                num nValue[3]
            mdesc mMdesc = {accel=25, vel=50, leave=1}
            num nActionIndex = 8
            num nDelay
            num nMoveType = 1
            num nPercentage
            num nSigValue = 1
        pointRx pPointRx[2] = {x=594.549716, y=30.77075, z=284.629716, rx=-40.404847, ry=94.502137, rz=40.914396, shoulder=lefty, elbow=epositive, wrist=wnegative}
        string sID
      [17]
        bool bMarked
        jointRx jJointRx = {j1=-1.639045, j2=12.402747, j3=111.595585, j4=2.517874, j5=-30.594648, j6=-1.669011}
        pointRx pInter
        paraItem pParaItem
          [0]
            bool bSafePoint
            ifItem iIfItem
              [0]
                bool bANDOR[2]
                num nSigIndex[3]
                num nSigType[3]
                num nValue[3]
            mdesc mMdesc
            num nActionIndex = 10
            num nDelay = 5
            num nMoveType = 4
            num nPercentage
            num nSigValue
        pointRx pPointRx[2] = {x=594.549819, y=30.770866, z=171.45682, rx=-40.410864, ry=94.502866, rz=40.920287, shoulder=lefty, elbow=epositive, wrist=wnegative}
        string sID
      [18]
        bool bMarked
        jointRx jJointRx = {j1=-1.639045, j2=12.402747, j3=111.595585, j4=2.517874, j5=-30.594648, j6=-1.669011}
        pointRx pInter
        paraItem pParaItem
          [0]
            bool bSafePoint
            ifItem iIfItem
              [0]
                bool bANDOR[2]
                num nSigIndex[3]
                num nSigType[3]
                num nValue[3]
            mdesc mMdesc
            num nActionIndex = 10
            num nDelay = 0.5
            num nMoveType = 7
            num nPercentage
            num nSigValue
        pointRx pPointRx[2] = {x=594.549819, y=30.770866, z=171.45682, rx=-40.410864, ry=94.502866, rz=40.920287, shoulder=lefty, elbow=epositive, wrist=wnegative}
        string sID
      [19]
        bool bMarked
        jointRx jJointRx = {j1=-1.639045, j2=12.402747, j3=111.595585, j4=2.517874, j5=-30.594648, j6=-1.669011}
        pointRx pInter
        paraItem pParaItem
          [0]
            bool bSafePoint
            ifItem iIfItem
              [0]
                bool bANDOR[2]
                num nSigIndex[3]
                num nSigType[3]
                num nValue[3]
            mdesc mMdesc
            num nActionIndex = 9
            num nDelay = 5
            num nMoveType = 3
            num nPercentage
            num nSigValue = 1
        pointRx pPointRx[2] = {x=594.549819, y=30.770866, z=171.45682, rx=-40.410864, ry=94.502866, rz=40.920287, shoulder=lefty, elbow=epositive, wrist=wnegative}
        string sID
      [20]
        bool bMarked
        jointRx jJointRx = {j1=-1.639045, j2=12.402747, j3=111.595585, j4=2.517874, j5=-30.594648, j6=-1.669011}
        pointRx pInter
        paraItem pParaItem
          [0]
            bool bSafePoint
            ifItem iIfItem
              [0]
                bool bANDOR[2]
                num nSigIndex[3]
                num nSigType[3]
                num nValue[3]
            mdesc mMdesc
            num nActionIndex = 9
            num nDelay = 5
            num nMoveType
            num nPercentage
            num nSigValue = 1
        pointRx pPointRx[2] = {x=594.549819, y=30.770866, z=171.45682, rx=-40.410864, ry=94.502866, rz=40.920287, shoulder=lefty, elbow=epositive, wrist=wnegative}
        string sID
      [21]
        bool bMarked
        jointRx jJointRx = {j1=-1.639045, j2=12.402747, j3=111.595585, j4=2.517874, j5=-30.594648, j6=-1.669011}
        pointRx pInter
        paraItem pParaItem
          [0]
            bool bSafePoint
            ifItem iIfItem
              [0]
                bool bANDOR[2]
                num nSigIndex[3]
                num nSigType[3]
                num nValue[3]
            mdesc mMdesc
            num nActionIndex = 9
            num nDelay = 5
            num nMoveType = 1
            num nPercentage
            num nSigValue = 1
        pointRx pPointRx[2] = {x=594.549819, y=30.770866, z=171.45682, rx=-40.410864, ry=94.502866, rz=40.920287, shoulder=lefty, elbow=epositive, wrist=wnegative}
        string sID
      [22]
        bool bMarked
        jointRx jJointRx = {j1=-1.639045, j2=12.402747, j3=111.595585, j4=2.517874, j5=-30.594648, j6=-1.669011}
        pointRx pInter
        paraItem pParaItem
          [0]
            bool bSafePoint
            ifItem iIfItem
              [0]
                bool bANDOR[2]
                num nSigIndex[3]
                num nSigType[3]
                num nValue[3]
            mdesc mMdesc
            num nActionIndex = 1
            num nDelay = 5
            num nMoveType = 6
            num nPercentage
            num nSigValue = 3
        pointRx pPointRx[2] = {x=594.549819, y=30.770866, z=171.45682, rx=-40.410864, ry=94.502866, rz=40.920287, shoulder=lefty, elbow=epositive, wrist=wnegative}
        string sID
      [23]
        bool bMarked
        jointRx jJointRx = {j1=-1.639045, j2=12.402747, j3=111.595585, j4=2.517874, j5=-30.594648, j6=-1.669011}
        pointRx pInter
        paraItem pParaItem
          [0]
            bool bSafePoint
            ifItem iIfItem
              [0]
                bool bANDOR[2]
                num nSigIndex[3]
                num nSigType[3]
                num nValue[3]
            mdesc mMdesc
            num nActionIndex = 1
            num nDelay = 5
            num nMoveType = 5
            num nPercentage
            num nSigValue = 3
        pointRx pPointRx[2] = {x=594.549819, y=30.770866, z=171.45682, rx=-40.410864, ry=94.502866, rz=40.920287, shoulder=lefty, elbow=epositive, wrist=wnegative}
        string sID
      [24]
        bool bMarked
        jointRx jJointRx = {j1=-1.639045, j2=12.402747, j3=111.595585, j4=2.517874, j5=-30.594648, j6=-1.669011}
        pointRx pInter
        paraItem pParaItem
          [0]
            bool bSafePoint
            ifItem iIfItem
              [0]
                bool bANDOR[2]
                num nSigIndex[3]
                num nSigType[3]
                num nValue[3]
            mdesc mMdesc
            num nActionIndex = 10
            num nDelay
            num nMoveType = 4
            num nPercentage
            num nSigValue = 1
        pointRx pPointRx[2] = {x=594.549819, y=30.770866, z=171.45682, rx=-40.410864, ry=94.502866, rz=40.920287, shoulder=lefty, elbow=epositive, wrist=wnegative}
        string sID
      [25]
        bool bMarked
        jointRx jJointRx = {j1=-1.639045, j2=12.402747, j3=111.595585, j4=2.517874, j5=-30.594648, j6=-1.669011}
        pointRx pInter
        paraItem pParaItem
          [0]
            bool bSafePoint
            ifItem iIfItem
              [0]
                bool bANDOR[2]
                num nSigIndex[3]
                num nSigType[3]
                num nValue[3]
            mdesc mMdesc
            num nActionIndex = 8
            num nDelay
            num nMoveType = 3
            num nPercentage
            num nSigValue = 1
        pointRx pPointRx[2] = {x=594.549819, y=30.770866, z=171.45682, rx=-40.410864, ry=94.502866, rz=40.920287, shoulder=lefty, elbow=epositive, wrist=wnegative}
        string sID
      [26]
        bool bMarked
        jointRx jJointRx = {j1=-1.639134, j2=22.193742, j3=116.03978, j4=1.817031, j5=-44.819098, j6=-0.790246}
        pointRx pInter
        paraItem pParaItem
          [0]
            bool bSafePoint
            ifItem iIfItem
              [0]
                bool bANDOR[2]
                num nSigIndex[3]
                num nSigType[3]
                num nValue[3]
            mdesc mMdesc = {accel=25, vel=50, leave=1}
            num nActionIndex = 8
            num nDelay
            num nMoveType = 1
            num nPercentage
            num nSigValue = 1
        pointRx pPointRx[2] = {x=594.549757, y=30.770873, z=70.540177, rx=-40.399083, ry=94.503271, rz=40.908669, shoulder=lefty, elbow=epositive, wrist=wnegative}
        string sID
      [27]
        bool bMarked
        jointRx jJointRx = {j1=-1.639045, j2=12.402747, j3=111.595585, j4=2.517874, j5=-30.594648, j6=-1.669011}
        pointRx pInter
        paraItem pParaItem
          [0]
            bool bSafePoint
            ifItem iIfItem
              [0]
                bool bANDOR[2]
                num nSigIndex[3]
                num nSigType[3]
                num nValue[3]
            mdesc mMdesc
            num nActionIndex = 10
            num nDelay = 5
            num nMoveType = 4
            num nPercentage
            num nSigValue
        pointRx pPointRx[2] = {x=594.549819, y=30.770866, z=171.45682, rx=-40.410864, ry=94.502866, rz=40.920287, shoulder=lefty, elbow=epositive, wrist=wnegative}
        string sID
      [28]
        bool bMarked
        jointRx jJointRx = {j1=-1.639045, j2=12.402747, j3=111.595585, j4=2.517874, j5=-30.594648, j6=-1.669011}
        pointRx pInter
        paraItem pParaItem
          [0]
            bool bSafePoint
            ifItem iIfItem
              [0]
                bool bANDOR[2]
                num nSigIndex[3]
                num nSigType[3]
                num nValue[3]
            mdesc mMdesc
            num nActionIndex = 10
            num nDelay = 0.5
            num nMoveType = 7
            num nPercentage
            num nSigValue
        pointRx pPointRx[2] = {x=594.549819, y=30.770866, z=171.45682, rx=-40.410864, ry=94.502866, rz=40.920287, shoulder=lefty, elbow=epositive, wrist=wnegative}
        string sID
      [29]
        bool bMarked
        jointRx jJointRx = {j1=-1.639045, j2=12.402747, j3=111.595585, j4=2.517874, j5=-30.594648, j6=-1.669011}
        pointRx pInter
        paraItem pParaItem
          [0]
            bool bSafePoint
            ifItem iIfItem
              [0]
                bool bANDOR[2]
                num nSigIndex[3]
                num nSigType[3]
                num nValue[3]
            mdesc mMdesc
            num nActionIndex = 9
            num nDelay = 5
            num nMoveType = 3
            num nPercentage
            num nSigValue = 1
        pointRx pPointRx[2] = {x=594.549819, y=30.770866, z=171.45682, rx=-40.410864, ry=94.502866, rz=40.920287, shoulder=lefty, elbow=epositive, wrist=wnegative}
        string sID
      [30]
        bool bMarked
        jointRx jJointRx = {j1=-1.639045, j2=12.402747, j3=111.595585, j4=2.517874, j5=-30.594648, j6=-1.669011}
        pointRx pInter
        paraItem pParaItem
          [0]
            bool bSafePoint
            ifItem iIfItem
              [0]
                bool bANDOR[2]
                num nSigIndex[3]
                num nSigType[3]
                num nValue[3]
            mdesc mMdesc
            num nActionIndex = 1
            num nDelay = 5
            num nMoveType = 6
            num nPercentage
            num nSigValue
        pointRx pPointRx[2] = {x=594.549819, y=30.770866, z=171.45682, rx=-40.410864, ry=94.502866, rz=40.920287, shoulder=lefty, elbow=epositive, wrist=wnegative}
        string sID
      [31]
        bool bMarked
        jointRx jJointRx = {j1=-1.639045, j2=12.402747, j3=111.595585, j4=2.517874, j5=-30.594648, j6=-1.669011}
        pointRx pInter
        paraItem pParaItem
          [0]
            bool bSafePoint
            ifItem iIfItem
              [0]
                bool bANDOR[2]
                num nSigIndex[3]
                num nSigType[3]
                num nValue[3]
            mdesc mMdesc
            num nActionIndex = 1
            num nDelay = 5
            num nMoveType = 5
            num nPercentage
            num nSigValue
        pointRx pPointRx[2] = {x=594.549819, y=30.770866, z=171.45682, rx=-40.410864, ry=94.502866, rz=40.920287, shoulder=lefty, elbow=epositive, wrist=wnegative}
        string sID
      [32]
        bool bMarked
        jointRx jJointRx = {j1=-6.64887, j2=-3.725236, j3=129.0447824, j4=-6.346176, j5=-34.648626, j6=4.794545}
        pointRx pInter
        paraItem pParaItem
          [0]
            bool bSafePoint
            ifItem iIfItem
              [0]
                bool bANDOR[2]
                num nSigIndex[3]
                num nSigType[3]
                num nValue[3]
            mdesc mMdesc
            num nActionIndex = 1
            num nDelay = 5
            num nMoveType
            num nPercentage
            num nSigValue
        pointRx pPointRx[2] = {x=472.316216, y=1.60837, z=176.938996, rx=-74.680282, ry=93.157396, rz=74.321891, shoulder=lefty, elbow=epositive, wrist=wnegative}
        string sID
      [33]
        bool bMarked
        jointRx jJointRx = {j1=-1.639045, j2=12.402747, j3=111.595585, j4=2.517874, j5=-30.594648, j6=-1.669011}
        pointRx pInter
        paraItem pParaItem
          [0]
            bool bSafePoint
            ifItem iIfItem
              [0]
                bool bANDOR[2]
                num nSigIndex[3]
                num nSigType[3]
                num nValue[3]
            mdesc mMdesc
            num nActionIndex = 11
            num nDelay = 5
            num nMoveType = 4
            num nPercentage
            num nSigValue = 1
        pointRx pPointRx[2] = {x=594.549819, y=30.770866, z=171.45682, rx=-40.410864, ry=94.502866, rz=40.920287, shoulder=lefty, elbow=epositive, wrist=wnegative}
        string sID
      [34]
        bool bMarked
        jointRx jJointRx = {j1=-1.639045, j2=12.402747, j3=111.595585, j4=2.517874, j5=-30.594648, j6=-1.669011}
        pointRx pInter
        paraItem pParaItem
          [0]
            bool bSafePoint
            ifItem iIfItem
              [0]
                bool bANDOR[2]
                num nSigIndex[3]
                num nSigType[3]
                num nValue[3]
            mdesc mMdesc
            num nActionIndex = 10
            num nDelay = 5
            num nMoveType = 3
            num nPercentage
            num nSigValue
        pointRx pPointRx[2] = {x=594.549819, y=30.770866, z=171.45682, rx=-40.410864, ry=94.502866, rz=40.920287, shoulder=lefty, elbow=epositive, wrist=wnegative}
        string sID
      [35]
        bool bMarked
        jointRx jJointRx = {j1=-1.639045, j2=12.402747, j3=111.595585, j4=2.517874, j5=-30.594648, j6=-1.669011}
        pointRx pInter
        paraItem pParaItem
          [0]
            bool bSafePoint
            ifItem iIfItem
              [0]
                bool bANDOR[2]
                num nSigIndex[3]
                num nSigType[3]
                num nValue[3]
            mdesc mMdesc
            num nActionIndex = 9
            num nDelay = 5
            num nMoveType = 4
            num nPercentage
            num nSigValue
        pointRx pPointRx[2] = {x=594.549819, y=30.770866, z=171.45682, rx=-40.410864, ry=94.502866, rz=40.920287, shoulder=lefty, elbow=epositive, wrist=wnegative}
        string sID
      [36]
        bool bMarked
        jointRx jJointRx = {j1=-1.639045, j2=12.402747, j3=111.595585, j4=2.517874, j5=-30.594648, j6=-1.669011}
        pointRx pInter
        paraItem pParaItem
          [0]
            bool bSafePoint
            ifItem iIfItem
              [0]
                bool bANDOR[2]
                num nSigIndex[3]
                num nSigType[3]
                num nValue[3]
            mdesc mMdesc
            num nActionIndex = 11
            num nDelay = 5
            num nMoveType = 4
            num nPercentage
            num nSigValue
        pointRx pPointRx[2] = {x=594.549819, y=30.770866, z=171.45682, rx=-40.410864, ry=94.502866, rz=40.920287, shoulder=lefty, elbow=epositive, wrist=wnegative}
        string sID
    string sID
  [03 543-7-0741]
    num nFrameIndex
    num nMoveID
    num nToolIndex
    pointItem pPointItem[45]
      [0]
        bool bMarked
        jointRx jJointRx = {j1=-2.594987, j2=-12.391258, j3=136.392534, j4=0.644488, j5=-30.575639, j6=-0.113504}
        pointRx pInter
        paraItem pParaItem
          [0]
            bool bSafePoint
            ifItem iIfItem
              [0]
                bool bANDOR[2]
                num nSigIndex[3]
                num nSigType[3]
                num nValue[3]
            mdesc mMdesc
            num nActionIndex = 11
            num nDelay
            num nMoveType = 4
            num nPercentage
            num nSigValue
        pointRx pPointRx[2] = {x=412.772469, y=30.77087, z=171.456836, rx=-40.418431, ry=94.503508, rz=40.927655, shoulder=lefty, elbow=epositive, wrist=wnegative}
        string sID
      [1]
        bool bMarked
        jointRx jJointRx = {j1=-2.594987, j2=-12.391258, j3=136.392534, j4=0.644488, j5=-30.575639, j6=-0.113504}
        pointRx pInter
        paraItem pParaItem
          [0]
            bool bSafePoint
            ifItem iIfItem
              [0]
                bool bANDOR[2]
                num nSigIndex[3]
                num nSigType[3]
                num nValue[3]
            mdesc mMdesc
            num nActionIndex = 9
            num nDelay
            num nMoveType = 4
            num nPercentage
            num nSigValue = 1
        pointRx pPointRx[2] = {x=412.772469, y=30.77087, z=171.456836, rx=-40.418431, ry=94.503508, rz=40.927655, shoulder=lefty, elbow=epositive, wrist=wnegative}
        string sID
      [2]
        bool bMarked
        jointRx jJointRx = {j1=-6.652009, j2=-3.724795, j3=129.0452396, j4=-6.346388, j5=-34.648815, j6=4.794651}
        pointRx pInter
        paraItem pParaItem
          [0]
            bool bSafePoint
            ifItem iIfItem
              [0]
                bool bANDOR[2]
                num nSigIndex[3]
                num nSigType[3]
                num nValue[3]
            mdesc mMdesc
            num nActionIndex = 9
            num nDelay
            num nMoveType
            num nPercentage
            num nSigValue = 1
        pointRx pPointRx[2] = {x=472.315715, y=1.582801, z=176.932517, rx=-74.682061, ry=93.16048, rz=74.323701, shoulder=lefty, elbow=epositive, wrist=wnegative}
        string sID
      [3]
        bool bMarked
        jointRx jJointRx = {j1=-5.216696, j2=41.157983, j3=119.687087, j4=-3.870543, j5=-83.639221, j6=1.741467}
        pointRx pInter
        paraItem pParaItem
          [0]
            bool bSafePoint
            ifItem iIfItem
              [0]
                bool bANDOR[2]
                num nSigIndex[3]
                num nSigType[3]
                num nValue[3]
            mdesc mMdesc = {leave=0}
            num nActionIndex
            num nDelay
            num nMoveType
            num nPercentage
            num nSigValue
        pointRx pPointRx[2] = {x=569.273857, y=4.969303, z=-59.417719, rx=5.605502, ry=77.187242, rz=-5.307477, shoulder=lefty, elbow=epositive, wrist=wnegative}
        string sID
      [4]
        bool bMarked
        jointRx jJointRx = {j1=-1.639045, j2=12.402747, j3=111.595585, j4=2.517874, j5=-30.594648, j6=-1.669011}
        pointRx pInter
        paraItem pParaItem
          [0]
            bool bSafePoint
            ifItem iIfItem
              [0]
                bool bANDOR[2]
                num nSigIndex[3]
                num nSigType[3]
                num nValue[3]
            mdesc mMdesc
            num nActionIndex = 1
            num nDelay
            num nMoveType = 6
            num nPercentage
            num nSigValue = 1
        pointRx pPointRx[2] = {x=594.549819, y=30.770866, z=171.45682, rx=-40.410864, ry=94.502866, rz=40.920287, shoulder=lefty, elbow=epositive, wrist=wnegative}
        string sID
      [5]
        bool bMarked
        jointRx jJointRx = {j1=-1.639045, j2=12.402747, j3=111.595585, j4=2.517874, j5=-30.594648, j6=-1.669011}
        pointRx pInter
        paraItem pParaItem
          [0]
            bool bSafePoint
            ifItem iIfItem
              [0]
                bool bANDOR[2]
                num nSigIndex[3]
                num nSigType[3]
                num nValue[3]
            mdesc mMdesc
            num nActionIndex = 1
            num nDelay
            num nMoveType = 5
            num nPercentage
            num nSigValue = 1
        pointRx pPointRx[2] = {x=594.549819, y=30.770866, z=171.45682, rx=-40.410864, ry=94.502866, rz=40.920287, shoulder=lefty, elbow=epositive, wrist=wnegative}
        string sID
      [6]
        bool bMarked
        jointRx jJointRx = {j1=-1.639045, j2=12.402747, j3=111.595585, j4=2.517874, j5=-30.594648, j6=-1.669011}
        pointRx pInter
        paraItem pParaItem
          [0]
            bool bSafePoint
            ifItem iIfItem
              [0]
                bool bANDOR[2]
                num nSigIndex[3]
                num nSigType[3]
                num nValue[3]
            mdesc mMdesc
            num nActionIndex = 10
            num nDelay
            num nMoveType = 4
            num nPercentage
            num nSigValue = 1
        pointRx pPointRx[2] = {x=594.549819, y=30.770866, z=171.45682, rx=-40.410864, ry=94.502866, rz=40.920287, shoulder=lefty, elbow=epositive, wrist=wnegative}
        string sID
      [7]
        bool bMarked
        jointRx jJointRx = {j1=-1.639045, j2=12.402747, j3=111.595585, j4=2.517874, j5=-30.594648, j6=-1.669011}
        pointRx pInter
        paraItem pParaItem
          [0]
            bool bSafePoint
            ifItem iIfItem
              [0]
                bool bANDOR[2]
                num nSigIndex[3]
                num nSigType[3]
                num nValue[3]
            mdesc mMdesc
            num nActionIndex = 8
            num nDelay
            num nMoveType = 3
            num nPercentage
            num nSigValue = 1
        pointRx pPointRx[2] = {x=594.549819, y=30.770866, z=171.45682, rx=-40.410864, ry=94.502866, rz=40.920287, shoulder=lefty, elbow=epositive, wrist=wnegative}
        string sID
      [8]
        bool bMarked
        jointRx jJointRx = {j1=-5.222925, j2=7.420427, j3=113.595368, j4=-5.551627, j5=-43.939511, j6=5.317784}
        pointRx pInter
        paraItem pParaItem
          [0]
            bool bSafePoint
            ifItem iIfItem
              [0]
                bool bANDOR[2]
                num nSigIndex[3]
                num nSigType[3]
                num nValue[3]
            mdesc mMdesc = {accel=0.64, vel=8, blend=cartesian, leave=0.1}
            num nActionIndex = 8
            num nDelay
            num nMoveType = 1
            num nPercentage
            num nSigValue = 1
        pointRx pPointRx[2] = {x=569.234173, y=4.915381, z=224.535515, rx=5.616876, ry=77.177601, rz=-5.318403, shoulder=lefty, elbow=epositive, wrist=wnegative}
        string sID
      [9]
        bool bMarked
        jointRx jJointRx = {j1=-1.639045, j2=12.402747, j3=111.595585, j4=2.517874, j5=-30.594648, j6=-1.669011}
        pointRx pInter
        paraItem pParaItem
          [0]
            bool bSafePoint
            ifItem iIfItem
              [0]
                bool bANDOR[2]
                num nSigIndex[3]
                num nSigType[3]
                num nValue[3]
            mdesc mMdesc
            num nActionIndex = 10
            num nDelay = 5
            num nMoveType = 4
            num nPercentage
            num nSigValue
        pointRx pPointRx[2] = {x=594.549819, y=30.770866, z=171.45682, rx=-40.410864, ry=94.502866, rz=40.920287, shoulder=lefty, elbow=epositive, wrist=wnegative}
        string sID
      [10]
        bool bMarked
        jointRx jJointRx = {j1=-1.639045, j2=12.402747, j3=111.595585, j4=2.517874, j5=-30.594648, j6=-1.669011}
        pointRx pInter
        paraItem pParaItem
          [0]
            bool bSafePoint
            ifItem iIfItem
              [0]
                bool bANDOR[2]
                num nSigIndex[3]
                num nSigType[3]
                num nValue[3]
            mdesc mMdesc
            num nActionIndex = 9
            num nDelay = 5
            num nMoveType = 3
            num nPercentage
            num nSigValue = 1
        pointRx pPointRx[2] = {x=594.549819, y=30.770866, z=171.45682, rx=-40.410864, ry=94.502866, rz=40.920287, shoulder=lefty, elbow=epositive, wrist=wnegative}
        string sID
      [11]
        bool bMarked
        jointRx jJointRx = {j1=-9.0335006, j2=-16.746462, j3=136.128627, j4=-8.563643, j5=-42.486188, j6=8.778813}
        pointRx pInter
        paraItem pParaItem
          [0]
            bool bSafePoint
            ifItem iIfItem
              [0]
                bool bANDOR[2]
                num nSigIndex[3]
                num nSigType[3]
                num nValue[3]
            mdesc mMdesc
            num nActionIndex
            num nDelay
            num nMoveType
            num nPercentage
            num nSigValue
        pointRx pPointRx[2] = {x=399.43075, y=-2.691352, z=220.472382, rx=13.539652, ry=76.911742, rz=-12.752112, shoulder=lefty, elbow=epositive, wrist=wnegative}
        string sID
      [12]
        bool bMarked
        jointRx jJointRx = {j1=-4.455815, j2=17.911136, j3=52.430951, j4=2.979533, j5=64.204099, j6=-3.394853}
        pointRx pInter
        paraItem pParaItem
          [0]
            bool bSafePoint
            ifItem iIfItem
              [0]
                bool bANDOR[2]
                num nSigIndex[3]
                num nSigType[3]
                num nValue[3]
            mdesc mMdesc
            num nActionIndex
            num nDelay
            num nMoveType
            num nPercentage
            num nSigValue
        pointRx pPointRx[2] = {x=654.439818, y=3.847964, z=477.339976, rx=-0.709996, ry=134.458429, rz=1.531981, shoulder=lefty, elbow=epositive, wrist=wpositive}
        string sID
      [13]
        bool bMarked
        jointRx jJointRx = {j1=-1.639045, j2=12.402747, j3=111.595585, j4=2.517874, j5=-30.594648, j6=-1.669011}
        pointRx pInter
        paraItem pParaItem
          [0]
            bool bSafePoint
            ifItem iIfItem
              [0]
                bool bANDOR[2]
                num nSigIndex[3]
                num nSigType[3]
                num nValue[3]
            mdesc mMdesc
            num nActionIndex = 1
            num nDelay
            num nMoveType = 6
            num nPercentage
            num nSigValue = 2
        pointRx pPointRx[2] = {x=594.549819, y=30.770866, z=171.45682, rx=-40.410864, ry=94.502866, rz=40.920287, shoulder=lefty, elbow=epositive, wrist=wnegative}
        string sID
      [14]
        bool bMarked
        jointRx jJointRx = {j1=-1.639045, j2=12.402747, j3=111.595585, j4=2.517874, j5=-30.594648, j6=-1.669011}
        pointRx pInter
        paraItem pParaItem
          [0]
            bool bSafePoint
            ifItem iIfItem
              [0]
                bool bANDOR[2]
                num nSigIndex[3]
                num nSigType[3]
                num nValue[3]
            mdesc mMdesc
            num nActionIndex = 1
            num nDelay
            num nMoveType = 5
            num nPercentage
            num nSigValue = 2
        pointRx pPointRx[2] = {x=594.549819, y=30.770866, z=171.45682, rx=-40.410864, ry=94.502866, rz=40.920287, shoulder=lefty, elbow=epositive, wrist=wnegative}
        string sID
      [15]
        bool bMarked
        jointRx jJointRx = {j1=-1.639045, j2=12.402747, j3=111.595585, j4=2.517874, j5=-30.594648, j6=-1.669011}
        pointRx pInter
        paraItem pParaItem
          [0]
            bool bSafePoint
            ifItem iIfItem
              [0]
                bool bANDOR[2]
                num nSigIndex[3]
                num nSigType[3]
                num nValue[3]
            mdesc mMdesc
            num nActionIndex = 10
            num nDelay
            num nMoveType = 4
            num nPercentage
            num nSigValue = 1
        pointRx pPointRx[2] = {x=594.549819, y=30.770866, z=171.45682, rx=-40.410864, ry=94.502866, rz=40.920287, shoulder=lefty, elbow=epositive, wrist=wnegative}
        string sID
      [16]
        bool bMarked
        jointRx jJointRx = {j1=-1.639045, j2=12.402747, j3=111.595585, j4=2.517874, j5=-30.594648, j6=-1.669011}
        pointRx pInter
        paraItem pParaItem
          [0]
            bool bSafePoint
            ifItem iIfItem
              [0]
                bool bANDOR[2]
                num nSigIndex[3]
                num nSigType[3]
                num nValue[3]
            mdesc mMdesc
            num nActionIndex = 8
            num nDelay
            num nMoveType = 3
            num nPercentage
            num nSigValue = 1
        pointRx pPointRx[2] = {x=594.549819, y=30.770866, z=171.45682, rx=-40.410864, ry=94.502866, rz=40.920287, shoulder=lefty, elbow=epositive, wrist=wnegative}
        string sID
      [17]
        bool bMarked
        jointRx jJointRx = {j1=-1.639045, j2=12.402747, j3=111.595585, j4=2.517874, j5=-30.594648, j6=-1.669011}
        pointRx pInter
        paraItem pParaItem
          [0]
            bool bSafePoint
            ifItem iIfItem
              [0]
                bool bANDOR[2]
                num nSigIndex[3]
                num nSigType[3]
                num nValue[3]
            mdesc mMdesc
            num nActionIndex = 8
            num nDelay
            num nMoveType = 7
            num nPercentage
            num nSigValue = 1
        pointRx pPointRx[2] = {x=594.549819, y=30.770866, z=171.45682, rx=-40.410864, ry=94.502866, rz=40.920287, shoulder=lefty, elbow=epositive, wrist=wnegative}
        string sID
      [18]
        bool bMarked
        jointRx jJointRx = {j1=-1.639045, j2=12.402747, j3=111.595585, j4=2.517874, j5=-30.594648, j6=-1.669011}
        pointRx pInter
        paraItem pParaItem
          [0]
            bool bSafePoint
            ifItem iIfItem
              [0]
                bool bANDOR[2]
                num nSigIndex[3]
                num nSigType[3]
                num nValue[3]
            mdesc mMdesc
            num nActionIndex = 10
            num nDelay = 5
            num nMoveType = 4
            num nPercentage
            num nSigValue
        pointRx pPointRx[2] = {x=594.549819, y=30.770866, z=171.45682, rx=-40.410864, ry=94.502866, rz=40.920287, shoulder=lefty, elbow=epositive, wrist=wnegative}
        string sID
      [19]
        bool bMarked
        jointRx jJointRx = {j1=-1.639045, j2=12.402747, j3=111.595585, j4=2.517874, j5=-30.594648, j6=-1.669011}
        pointRx pInter
        paraItem pParaItem
          [0]
            bool bSafePoint
            ifItem iIfItem
              [0]
                bool bANDOR[2]
                num nSigIndex[3]
                num nSigType[3]
                num nValue[3]
            mdesc mMdesc
            num nActionIndex = 10
            num nDelay = 0.5
            num nMoveType = 7
            num nPercentage
            num nSigValue
        pointRx pPointRx[2] = {x=594.549819, y=30.770866, z=171.45682, rx=-40.410864, ry=94.502866, rz=40.920287, shoulder=lefty, elbow=epositive, wrist=wnegative}
        string sID
      [20]
        bool bMarked
        jointRx jJointRx = {j1=-1.639045, j2=12.402747, j3=111.595585, j4=2.517874, j5=-30.594648, j6=-1.669011}
        pointRx pInter
        paraItem pParaItem
          [0]
            bool bSafePoint
            ifItem iIfItem
              [0]
                bool bANDOR[2]
                num nSigIndex[3]
                num nSigType[3]
                num nValue[3]
            mdesc mMdesc
            num nActionIndex = 9
            num nDelay = 5
            num nMoveType = 3
            num nPercentage
            num nSigValue = 1
        pointRx pPointRx[2] = {x=594.549819, y=30.770866, z=171.45682, rx=-40.410864, ry=94.502866, rz=40.920287, shoulder=lefty, elbow=epositive, wrist=wnegative}
        string sID
      [21]
        bool bMarked
        jointRx jJointRx = {j1=-4.814062, j2=18.435461, j3=46.904954, j4=3.142299, j5=69.216348, j6=-3.464711}
        pointRx pInter
        paraItem pParaItem
          [0]
            bool bSafePoint
            ifItem iIfItem
              [0]
                bool bANDOR[2]
                num nSigIndex[3]
                num nSigType[3]
                num nValue[3]
            mdesc mMdesc = {leave=0}
            num nActionIndex = 9
            num nDelay = 5
            num nMoveType
            num nPercentage
            num nSigValue = 1
        pointRx pPointRx[2] = {x=644.200475, y=1.0657947, z=510.476498, rx=-0.710255, ry=134.458452, rz=1.532258, shoulder=lefty, elbow=epositive, wrist=wpositive}
        string sID
      [22]
        bool bMarked
        jointRx jJointRx = {j1=-1.639045, j2=12.402747, j3=111.595585, j4=2.517874, j5=-30.594648, j6=-1.669011}
        pointRx pInter
        paraItem pParaItem
          [0]
            bool bSafePoint
            ifItem iIfItem
              [0]
                bool bANDOR[2]
                num nSigIndex[3]
                num nSigType[3]
                num nValue[3]
            mdesc mMdesc
            num nActionIndex = 1
            num nDelay = 5
            num nMoveType = 6
            num nPercentage
            num nSigValue = 3
        pointRx pPointRx[2] = {x=594.549819, y=30.770866, z=171.45682, rx=-40.410864, ry=94.502866, rz=40.920287, shoulder=lefty, elbow=epositive, wrist=wnegative}
        string sID
      [23]
        bool bMarked
        jointRx jJointRx = {j1=-1.639045, j2=12.402747, j3=111.595585, j4=2.517874, j5=-30.594648, j6=-1.669011}
        pointRx pInter
        paraItem pParaItem
          [0]
            bool bSafePoint
            ifItem iIfItem
              [0]
                bool bANDOR[2]
                num nSigIndex[3]
                num nSigType[3]
                num nValue[3]
            mdesc mMdesc
            num nActionIndex = 1
            num nDelay = 5
            num nMoveType = 5
            num nPercentage
            num nSigValue = 3
        pointRx pPointRx[2] = {x=594.549819, y=30.770866, z=171.45682, rx=-40.410864, ry=94.502866, rz=40.920287, shoulder=lefty, elbow=epositive, wrist=wnegative}
        string sID
      [24]
        bool bMarked
        jointRx jJointRx = {j1=-1.639045, j2=12.402747, j3=111.595585, j4=2.517874, j5=-30.594648, j6=-1.669011}
        pointRx pInter
        paraItem pParaItem
          [0]
            bool bSafePoint
            ifItem iIfItem
              [0]
                bool bANDOR[2]
                num nSigIndex[3]
                num nSigType[3]
                num nValue[3]
            mdesc mMdesc
            num nActionIndex = 10
            num nDelay
            num nMoveType = 4
            num nPercentage
            num nSigValue = 1
        pointRx pPointRx[2] = {x=594.549819, y=30.770866, z=171.45682, rx=-40.410864, ry=94.502866, rz=40.920287, shoulder=lefty, elbow=epositive, wrist=wnegative}
        string sID
      [25]
        bool bMarked
        jointRx jJointRx = {j1=-1.639045, j2=12.402747, j3=111.595585, j4=2.517874, j5=-30.594648, j6=-1.669011}
        pointRx pInter
        paraItem pParaItem
          [0]
            bool bSafePoint
            ifItem iIfItem
              [0]
                bool bANDOR[2]
                num nSigIndex[3]
                num nSigType[3]
                num nValue[3]
            mdesc mMdesc
            num nActionIndex = 8
            num nDelay
            num nMoveType = 3
            num nPercentage
            num nSigValue = 1
        pointRx pPointRx[2] = {x=594.549819, y=30.770866, z=171.45682, rx=-40.410864, ry=94.502866, rz=40.920287, shoulder=lefty, elbow=epositive, wrist=wnegative}
        string sID
      [26]
        bool bMarked
        jointRx jJointRx = {j1=-4.813626, j2=14.411965, j3=88.10628, j4=5.527501, j5=32.129903, j6=-7.0332281}
        pointRx pInter
        paraItem pParaItem
